Fanuc KAREL source: KD00048.KL

PROGRAM KD00048
%NOLOCKGROUP
%DEFGROUP = 1
VAR
  I: INTEGER
  J: INTEGER
  B: BOOLEAN
  R: REAL
  S: STRING[80]
  PTH: PATH
BEGIN
  MOVE ALONG PTH
END KD00048
